(* PLC project GeneratedProgram, SafePLC-Gen SafePLC-Gen Multimodal 1.0 *)
(* stored: creationDateTime 2026-04-25T13:41:59.797045Z *)

PROGRAM GeneratedProgram
  VAR
    TICSA_4750_03_Scaled : REAL;
    PICSA_4712_02_Scaled : REAL;
    PI_4712_01_Scaled : REAL;
    TICSA_4750_03_HH_SP : REAL;
    TICSA_4750_03_H_SP : REAL;
    TICSA_4750_03_L_SP : REAL;
    TICSA_4750_03_LL_SP : REAL;
    TICSA_4750_03_Deadband : REAL;
    PICSA_4712_02_HH_SP : REAL;
    PICSA_4712_02_H_SP : REAL;
    PICSA_4712_02_L_SP : REAL;
    PICSA_4712_02_LL_SP : REAL;
    PICSA_4712_02_Deadband : REAL;
    PI_4712_01_HH_SP : REAL;
    PI_4712_01_H_SP : REAL;
    PI_4712_01_L_SP : REAL;
    PI_4712_01_LL_SP : REAL;
    PI_4712_01_Deadband : REAL;
    TICSA_4750_03_H : BOOL;
    TICSA_4750_03_L : BOOL;
    TICSA_4750_03_HH_Set : BOOL;
    TICSA_4750_03_HH_Rst : BOOL;
    TICSA_4750_03_LL_Set : BOOL;
    TICSA_4750_03_LL_Rst : BOOL;
    TICSA_4750_03_HH_Latch : SR;
    TICSA_4750_03_LL_Latch : SR;
    TICSA_4750_03_HH_Ack : BOOL;
    TICSA_4750_03_LL_Ack : BOOL;
    PICSA_4712_02_H : BOOL;
    PICSA_4712_02_L : BOOL;
    PICSA_4712_02_HH_Set : BOOL;
    PICSA_4712_02_HH_Rst : BOOL;
    PICSA_4712_02_LL_Set : BOOL;
    PICSA_4712_02_LL_Rst : BOOL;
    PICSA_4712_02_HH_Latch : SR;
    PICSA_4712_02_LL_Latch : SR;
    PICSA_4712_02_HH_Ack : BOOL;
    PICSA_4712_02_LL_Ack : BOOL;
    PI_4712_01_H : BOOL;
    PI_4712_01_L : BOOL;
    PI_4712_01_HH_Set : BOOL;
    PI_4712_01_HH_Rst : BOOL;
    PI_4712_01_LL_Set : BOOL;
    PI_4712_01_LL_Rst : BOOL;
    PI_4712_01_HH_Latch : SR;
    PI_4712_01_LL_Latch : SR;
    PI_4712_01_HH_Ack : BOOL;
    PI_4712_01_LL_Ack : BOOL;
    LOOP_4750_03_TRIP : BOOL;
    LOOP_4712_02_TRIP : BOOL;
    LOOP_104_01_TRIP : BOOL;
    SAFE_STATE : BOOL;
    TICSA_4750_03_HH : BOOL;
    TICSA_4750_03_LL : BOOL;
    PICSA_4712_02_HH : BOOL;
    PICSA_4712_02_LL : BOOL;
    SV_104_01_HH : BOOL;
    SV_104_01_LL : BOOL;
    TICSA_4750_03_SP : REAL;
    TICSA_4750_03_Error : REAL;
    TICSA_4750_03_Integral : REAL;
    TICSA_4750_03_Kp : REAL;
    TICSA_4750_03_Ki : REAL;
    TICSA_4750_03_Output : REAL;
    PICSA_4712_02_SP : REAL;
    PICSA_4712_02_Error : REAL;
    PICSA_4712_02_Integral : REAL;
    PICSA_4712_02_Kp : REAL;
    PICSA_4712_02_Ki : REAL;
    PICSA_4712_02_Output : REAL;
    SV_104_01_Out : BOOL;
    CHK_75SA21_80_Out : BOOL;
    CHK_MNc_47125_Out : BOOL;
    ISOV_73KH12_25_1_Out : BOOL;
    ISOV_73KH12_25_2_Out : BOOL;
    ISOV_73KH12_50_1_Out : BOOL;
    ISOV_73KH12_50_2_Out : BOOL;
    ISOV_73KH12_50_3_Out : BOOL;
    ISOV_MNb_47121_Out : BOOL;
    ISOV_MNb_47122_Out : BOOL;
    ISOV_MNb_47123_Out : BOOL;
    ISOV_MNc_47124_Out : BOOL;
    ISOV_MNc_47125_73HG12_Out : BOOL;
    ISOV_MNc_47126_Out : BOOL;
    ISOV_MNc_47127_Out : BOOL;
    ISOV_WKa_47130_Out : BOOL;
    ISOV_WKa_47131_Out : BOOL;
    ISOV_QSa_47140_Out : BOOL;
    ISOV_QSb_47141_Out : BOOL;
    System_Alarm : BOOL;
    FirstScan : BOOL;
  END_VAR

            IF FirstScan THEN
    LOOP_4750_03_TRIP      := TRUE;
    LOOP_4712_02_TRIP      := TRUE;
    LOOP_104_01_TRIP       := TRUE;
    SAFE_STATE             := TRUE;
    TV_4750_03_Out         := 6554;
    PVA_4712_02_Out        := 6554;
    FC_HV_H_1007_inlet_Out := 6554;
    SV_104_01_Out          := FALSE;
    TICSA_4750_03_Integral := 0.0;
    PICSA_4712_02_Integral := 0.0;
    TICSA_4750_03_HH_Latch(S1 := FALSE, R := TRUE);
    TICSA_4750_03_LL_Latch(S1 := FALSE, R := TRUE);
    PICSA_4712_02_HH_Latch(S1 := FALSE, R := TRUE);
    PICSA_4712_02_LL_Latch(S1 := FALSE, R := TRUE);
    PI_4712_01_HH_Latch(S1 := FALSE, R := TRUE);
    PI_4712_01_LL_Latch(S1 := FALSE, R := TRUE);
    FirstScan := FALSE;
    RETURN;
END_IF;

TICSA_4750_03_Scaled := ((INT_TO_REAL(TICSA_4750_03_Raw) - 6554.0) / (32767.0 - 6554.0)) * 150.0;
PICSA_4712_02_Scaled := ((INT_TO_REAL(PICSA_4712_02_Raw) - 6554.0) / (32767.0 - 6554.0)) * 25.0;
PI_4712_01_Scaled    := ((INT_TO_REAL(PI_4712_01_Raw)    - 6554.0) / (32767.0 - 6554.0)) * 25.0;

TICSA_4750_03_HH := TICSA_4750_03_Scaled >= TICSA_4750_03_HH_SP;
TICSA_4750_03_LL := TICSA_4750_03_Scaled <= TICSA_4750_03_LL_SP;
PICSA_4712_02_HH := PICSA_4712_02_Scaled >= PICSA_4712_02_HH_SP;
PICSA_4712_02_LL := PICSA_4712_02_Scaled <= PICSA_4712_02_LL_SP;

IF TICSA_4750_03_HH OR TICSA_4750_03_LL THEN
    LOOP_4750_03_TRIP := TRUE;
ELSIF LOOP_4750_03_TRIP AND MANUAL_RESET AND NOT TICSA_4750_03_HH AND NOT TICSA_4750_03_LL THEN
    LOOP_4750_03_TRIP := FALSE;
END_IF;

IF PICSA_4712_02_HH OR PICSA_4712_02_LL THEN
    LOOP_4712_02_TRIP := TRUE;
ELSIF LOOP_4712_02_TRIP AND MANUAL_RESET AND NOT PICSA_4712_02_HH AND NOT PICSA_4712_02_LL THEN
    LOOP_4712_02_TRIP := FALSE;
END_IF;

IF SV_104_01_HH OR SV_104_01_LL THEN
    LOOP_104_01_TRIP := TRUE;
ELSIF LOOP_104_01_TRIP AND MANUAL_RESET AND NOT SV_104_01_HH AND NOT SV_104_01_LL THEN
    LOOP_104_01_TRIP := FALSE;
END_IF;

SAFE_STATE := ESTOP OR LOOP_4750_03_TRIP OR LOOP_4712_02_TRIP OR LOOP_104_01_TRIP;

IF TICSA_4750_03_Scaled >= TICSA_4750_03_HH_SP THEN
    TICSA_4750_03_HH_Set := TRUE;
ELSIF TICSA_4750_03_Scaled <= (TICSA_4750_03_HH_SP - TICSA_4750_03_Deadband) THEN
    TICSA_4750_03_HH_Set := FALSE;
END_IF;
TICSA_4750_03_HH_Rst := TICSA_4750_03_HH_Ack AND NOT TICSA_4750_03_HH_Set;
TICSA_4750_03_HH_Latch(S1 := TICSA_4750_03_HH_Set, R := TICSA_4750_03_HH_Rst);

IF TICSA_4750_03_Scaled <= TICSA_4750_03_LL_SP THEN
    TICSA_4750_03_LL_Set := TRUE;
ELSIF TICSA_4750_03_Scaled >= (TICSA_4750_03_LL_SP + TICSA_4750_03_Deadband) THEN
    TICSA_4750_03_LL_Set := FALSE;
END_IF;
TICSA_4750_03_LL_Rst := TICSA_4750_03_LL_Ack AND NOT TICSA_4750_03_LL_Set;
TICSA_4750_03_LL_Latch(S1 := TICSA_4750_03_LL_Set, R := TICSA_4750_03_LL_Rst);

IF TICSA_4750_03_Scaled >= TICSA_4750_03_H_SP THEN
    TICSA_4750_03_H := TRUE;
ELSIF TICSA_4750_03_Scaled <= (TICSA_4750_03_H_SP - TICSA_4750_03_Deadband) THEN
    TICSA_4750_03_H := FALSE;
END_IF;

IF TICSA_4750_03_Scaled <= TICSA_4750_03_L_SP THEN
    TICSA_4750_03_L := TRUE;
ELSIF TICSA_4750_03_Scaled >= (TICSA_4750_03_L_SP + TICSA_4750_03_Deadband) THEN
    TICSA_4750_03_L := FALSE;
END_IF;

IF PICSA_4712_02_Scaled >= PICSA_4712_02_HH_SP THEN
    PICSA_4712_02_HH_Set := TRUE;
ELSIF PICSA_4712_02_Scaled <= (PICSA_4712_02_HH_SP - PICSA_4712_02_Deadband) THEN
    PICSA_4712_02_HH_Set := FALSE;
END_IF;
PICSA_4712_02_HH_Rst := PICSA_4712_02_HH_Ack AND NOT PICSA_4712_02_HH_Set;
PICSA_4712_02_HH_Latch(S1 := PICSA_4712_02_HH_Set, R := PICSA_4712_02_HH_Rst);

IF PICSA_4712_02_Scaled <= PICSA_4712_02_LL_SP THEN
    PICSA_4712_02_LL_Set := TRUE;
ELSIF PICSA_4712_02_Scaled >= (PICSA_4712_02_LL_SP + PICSA_4712_02_Deadband) THEN
    PICSA_4712_02_LL_Set := FALSE;
END_IF;
PICSA_4712_02_LL_Rst := PICSA_4712_02_LL_Ack AND NOT PICSA_4712_02_LL_Set;
PICSA_4712_02_LL_Latch(S1 := PICSA_4712_02_LL_Set, R := PICSA_4712_02_LL_Rst);

IF PICSA_4712_02_Scaled >= PICSA_4712_02_H_SP THEN
    PICSA_4712_02_H := TRUE;
ELSIF PICSA_4712_02_Scaled <= (PICSA_4712_02_H_SP - PICSA_4712_02_Deadband) THEN
    PICSA_4712_02_H := FALSE;
END_IF;

IF PICSA_4712_02_Scaled <= PICSA_4712_02_L_SP THEN
    PICSA_4712_02_L := TRUE;
ELSIF PICSA_4712_02_Scaled >= (PICSA_4712_02_L_SP + PICSA_4712_02_Deadband) THEN
    PICSA_4712_02_L := FALSE;
END_IF;

IF PI_4712_01_Scaled >= PI_4712_01_HH_SP THEN
    PI_4712_01_HH_Set := TRUE;
ELSIF PI_4712_01_Scaled <= (PI_4712_01_HH_SP - PI_4712_01_Deadband) THEN
    PI_4712_01_HH_Set := FALSE;
END_IF;
PI_4712_01_HH_Rst := PI_4712_01_HH_Ack AND NOT PI_4712_01_HH_Set;
PI_4712_01_HH_Latch(S1 := PI_4712_01_HH_Set, R := PI_4712_01_HH_Rst);

IF PI_4712_01_Scaled <= PI_4712_01_LL_SP THEN
    PI_4712_01_LL_Set := TRUE;
ELSIF PI_4712_01_Scaled >= (PI_4712_01_LL_SP + PI_4712_01_Deadband) THEN
    PI_4712_01_LL_Set := FALSE;
END_IF;
PI_4712_01_LL_Rst := PI_4712_01_LL_Ack AND NOT PI_4712_01_LL_Set;
PI_4712_01_LL_Latch(S1 := PI_4712_01_LL_Set, R := PI_4712_01_LL_Rst);

IF PI_4712_01_Scaled >= PI_4712_01_H_SP THEN
    PI_4712_01_H := TRUE;
ELSIF PI_4712_01_Scaled <= (PI_4712_01_H_SP - PI_4712_01_Deadband) THEN
    PI_4712_01_H := FALSE;
END_IF;

IF PI_4712_01_Scaled <= PI_4712_01_L_SP THEN
    PI_4712_01_L := TRUE;
ELSIF PI_4712_01_Scaled >= (PI_4712_01_L_SP + PI_4712_01_Deadband) THEN
    PI_4712_01_L := FALSE;
END_IF;

IF NOT SAFE_STATE THEN
    TICSA_4750_03_Error    := TICSA_4750_03_SP - TICSA_4750_03_Scaled;
    TICSA_4750_03_Integral := TICSA_4750_03_Integral + (TICSA_4750_03_Ki * TICSA_4750_03_Error);
    IF TICSA_4750_03_Integral > 100.0 THEN
        TICSA_4750_03_Integral := 100.0;
    ELSIF TICSA_4750_03_Integral < 0.0 THEN
        TICSA_4750_03_Integral := 0.0;
    END_IF;
    TICSA_4750_03_Output := (TICSA_4750_03_Kp * TICSA_4750_03_Error) + TICSA_4750_03_Integral;
    IF TICSA_4750_03_Output > 100.0 THEN
        TICSA_4750_03_Output := 100.0;
    ELSIF TICSA_4750_03_Output < 0.0 THEN
        TICSA_4750_03_Output := 0.0;
    END_IF;
    TV_4750_03_Out := REAL_TO_INT(6554.0 + (TICSA_4750_03_Output / 100.0) * (32767.0 - 6554.0));

    PICSA_4712_02_Error    := PICSA_4712_02_SP - PICSA_4712_02_Scaled;
    PICSA_4712_02_Integral := PICSA_4712_02_Integral + (PICSA_4712_02_Ki * PICSA_4712_02_Error);
    IF PICSA_4712_02_Integral > 100.0 THEN
        PICSA_4712_02_Integral := 100.0;
    ELSIF PICSA_4712_02_Integral < 0.0 THEN
        PICSA_4712_02_Integral := 0.0;
    END_IF;
    PICSA_4712_02_Output := (PICSA_4712_02_Kp * PICSA_4712_02_Error) + PICSA_4712_02_Integral;
    IF PICSA_4712_02_Output > 100.0 THEN
        PICSA_4712_02_Output := 100.0;
    ELSIF PICSA_4712_02_Output < 0.0 THEN
        PICSA_4712_02_Output := 0.0;
    END_IF;
    PVA_4712_02_Out := REAL_TO_INT(6554.0 + (PICSA_4712_02_Output / 100.0) * (32767.0 - 6554.0));

    IF HS_4750_01 THEN
        FC_HV_H_1007_inlet_Out := 32767;
    ELSE
        FC_HV_H_1007_inlet_Out := 6554;
    END_IF;

    SV_104_01_Out              := TRUE;
    CHK_75SA21_80_Out          := TRUE;
    CHK_MNc_47125_Out          := TRUE;
    ISOV_73KH12_25_1_Out       := TRUE;
    ISOV_73KH12_25_2_Out       := TRUE;
    ISOV_73KH12_50_1_Out       := TRUE;
    ISOV_73KH12_50_2_Out       := TRUE;
    ISOV_73KH12_50_3_Out       := TRUE;
    ISOV_MNb_47121_Out         := TRUE;
    ISOV_MNb_47122_Out         := TRUE;
    ISOV_MNb_47123_Out         := TRUE;
    ISOV_MNc_47124_Out         := TRUE;
    ISOV_MNc_47125_73HG12_Out  := TRUE;
    ISOV_MNc_47126_Out         := TRUE;
    ISOV_MNc_47127_Out         := TRUE;
    ISOV_WKa_47130_Out         := TRUE;
    ISOV_WKa_47131_Out         := TRUE;
    ISOV_QSa_47140_Out         := TRUE;
    ISOV_QSb_47141_Out         := TRUE;
ELSE
    TV_4750_03_Out             := 6554;
    PVA_4712_02_Out            := 6554;
    FC_HV_H_1007_inlet_Out     := 6554;
    SV_104_01_Out              := FALSE;
    CHK_75SA21_80_Out          := FALSE;
    CHK_MNc_47125_Out          := FALSE;
    ISOV_73KH12_25_1_Out       := FALSE;
    ISOV_73KH12_25_2_Out       := FALSE;
    ISOV_73KH12_50_1_Out       := FALSE;
    ISOV_73KH12_50_2_Out       := FALSE;
    ISOV_73KH12_50_3_Out       := FALSE;
    ISOV_MNb_47121_Out         := FALSE;
    ISOV_MNb_47122_Out         := FALSE;
    ISOV_MNb_47123_Out         := FALSE;
    ISOV_MNc_47124_Out         := FALSE;
    ISOV_MNc_47125_73HG12_Out  := FALSE;
    ISOV_MNc_47126_Out         := FALSE;
    ISOV_MNc_47127_Out         := FALSE;
    ISOV_WKa_47130_Out         := FALSE;
    ISOV_WKa_47131_Out         := FALSE;
    ISOV_QSa_47140_Out         := FALSE;
    ISOV_QSb_47141_Out         := FALSE;
END_IF;

System_Alarm :=
    TICSA_4750_03_HH_Latch.Q1 OR TICSA_4750_03_LL_Latch.Q1 OR
    TICSA_4750_03_H            OR TICSA_4750_03_L            OR
    PICSA_4712_02_HH_Latch.Q1 OR PICSA_4712_02_LL_Latch.Q1 OR
    PICSA_4712_02_H            OR PICSA_4712_02_L            OR
    PI_4712_01_HH_Latch.Q1    OR PI_4712_01_LL_Latch.Q1    OR
    PI_4712_01_H               OR PI_4712_01_L              OR
    LOOP_4750_03_TRIP          OR LOOP_4712_02_TRIP         OR
    LOOP_104_01_TRIP           OR ESTOP;
          
END_PROGRAM

CONFIGURATION Config0
  RESOURCE Res0 ON PLC
    TASK MainTask(INTERVAL := T#20ms, PRIORITY := 0);
    PROGRAM Main : GeneratedProgram;
  END_RESOURCE
END_CONFIGURATION
